// TIA Portal V21 program export: 0 tag tables, 0 data types, 1 data blocks, 1 code blocks (in call order from the OBs), 0 instance data blocks

DATA_BLOCK "DB_FAT_Demo"   // DB1
{ S7_Optimized_Access := 'FALSE' }
VERSION : 1.0
// SPDX-License-Identifier: MIT. Public passive laboratory example.
// stored: AutoNumber true, CodeModifiedDate 2026-11-03T19:44:32.7091278Z, CompileDate 2026-11-03T19:44:33.4739621Z, CreationDate 2026-11-03T19:44:31.2051572Z, DBAccessibleFromOPCUA true, DBAccessibleFromWebserver true, DownloadDate 0001-01-01T00:00:00Z, InterfaceModifiedDate 2026-11-03T19:44:32.7091278Z, IsConsistent true, IsKnowHowProtected false, IsOnlyStoredInLoadMemory false, IsPLCDB false, IsWriteProtectedInAS false, LoadMemoryLength 5286, ModifiedDate 2026-11-03T19:44:32.7091278Z, ParameterModified 2026-11-03T19:44:32.7091278Z, StructureModified 2026-11-03T19:44:32.7091278Z, WorkMemoryLength 192
   VAR RETAIN
      EnableDemo { ExternalAccessible := 'False'; ExternalVisible := 'False'; ExternalWritable := 'False'} : Bool := TRUE;   // isolated virtual copy only
      StopHealthy : Bool := TRUE;
      P101_Request : Bool := FALSE;
      P101_RequestedSpeed : Real := REAL#60.0;
      P101_RunCommand { ExternalWritable := 'False'} : Bool := FALSE;
      P101_SpeedCommand { ExternalWritable := 'False'} : Real := REAL#0.0;
      P101_Running : Bool := FALSE;
      P101_SpeedFeedback : Real := REAL#0.0;
      P101_Fault : Bool := FALSE;
      P201_Request : Bool := FALSE;
      P201_RequestedSpeed : Real := REAL#60.0;
      P201_RunCommand { ExternalWritable := 'False'} : Bool := FALSE;
      P201_SpeedCommand { ExternalWritable := 'False'} : Real := REAL#0.0;
      P201_Running : Bool := FALSE;
      P201_SpeedFeedback : Real := REAL#0.0;
      P201_Fault : Bool := FALSE;
      P202_Request : Bool := FALSE;
      P202_RequestedSpeed : Real := REAL#60.0;
      P202_RunCommand { ExternalWritable := 'False'} : Bool := FALSE;
      P202_SpeedCommand { ExternalWritable := 'False'} : Real := REAL#0.0;
      P202_Running : Bool := FALSE;
      P202_SpeedFeedback : Real := REAL#0.0;
      P202_Fault : Bool := FALSE;
      P301_Request : Bool := FALSE;
      P301_RequestedSpeed : Real := REAL#60.0;
      P301_RunCommand { ExternalWritable := 'False'} : Bool := FALSE;
      P301_SpeedCommand { ExternalWritable := 'False'} : Real := REAL#0.0;
      P301_Running : Bool := FALSE;
      P301_SpeedFeedback : Real := REAL#0.0;
      P301_Fault : Bool := FALSE;
      XV101_Request : Bool := FALSE;
      XV101_OpenCommand { ExternalWritable := 'False'} : Bool := FALSE;
      XV101_Open : Bool := FALSE;
      XV101_Closed : Bool := TRUE;
      XV201_Request : Bool := FALSE;
      XV201_OpenCommand { ExternalWritable := 'False'} : Bool := FALSE;
      XV201_Open : Bool := FALSE;
      XV201_Closed : Bool := TRUE;
      XV202_Request : Bool := FALSE;
      XV202_OpenCommand { ExternalWritable := 'False'} : Bool := FALSE;
      XV202_Open : Bool := FALSE;
      XV202_Closed : Bool := TRUE;
      XV301_Request : Bool := FALSE;
      XV301_OpenCommand { ExternalWritable := 'False'} : Bool := FALSE;
      XV301_Open : Bool := FALSE;
      XV301_Closed : Bool := TRUE;
      XV102_Request : Bool := FALSE;
      XV102_OpenCommand { ExternalWritable := 'False'} : Bool := FALSE;
      XV102_Open : Bool := FALSE;
      XV102_Closed : Bool := TRUE;
      XV203_Request : Bool := FALSE;
      XV203_OpenCommand { ExternalWritable := 'False'} : Bool := FALSE;
      XV203_Open : Bool := FALSE;
      XV203_Closed : Bool := TRUE;
      XV103_Request : Bool := FALSE;
      XV103_OpenCommand { ExternalWritable := 'False'} : Bool := FALSE;
      XV103_Open : Bool := FALSE;
      XV103_Closed : Bool := TRUE;
      FCV302_RequestedPosition : Real := REAL#0.0;
      FCV302_PositionCommand { ExternalWritable := 'False'} : Real := REAL#0.0;
      FCV302_PositionFeedback : Real := REAL#0.0;
      LT101_Raw : Int := INT#16589;
      LT101_Percent { ExternalWritable := 'False'} : Real := REAL#0.0;
      TK101_Volume : Real := REAL#720.0;
      LSL101 : Bool := FALSE;
      LSH101 : Bool := FALSE;
      LT201_Raw : Int := INT#6912;
      LT201_Percent { ExternalWritable := 'False'} : Real := REAL#0.0;
      TK201_Volume : Real := REAL#450.0;
      LSL201 : Bool := FALSE;
      LSH201 : Bool := FALSE;
      LT301_Raw : Int := INT#4147;
      LT301_Percent { ExternalWritable := 'False'} : Real := REAL#0.0;
      TK301_Volume : Real := REAL#180.0;
      LSL301 : Bool := FALSE;
      LSH301 : Bool := FALSE;
   END_VAR
BEGIN
END_DATA_BLOCK

ORGANIZATION_BLOCK "Main"   // OB1, SCL, ProgramCycle
{ S7_Optimized_Access := 'TRUE' }
VERSION : 1.0
// SPDX-License-Identifier: MIT. No equipment library or process sequence.
// stored: AutoNumber true, CodeModifiedDate 2026-11-03T19:44:43.8400479Z, CompileDate 2026-11-03T19:44:43.8400479Z, ConstantName OB_Main, CreationDate 2026-11-03T19:44:33.7000652Z, DownloadDate 0001-01-01T00:00:00Z, EventClass Program cycle, HandleErrorsWithinBlock false, InterfaceModifiedDate 2026-11-03T19:44:33.988557Z, IsConsistent true, IsIECCheckEnabled false, IsKnowHowProtected false, IsWriteProtected false, LoadMemoryLength 14729, ModifiedDate 2026-11-03T19:44:43.8400479Z, PLCSimAdvancedSupport true, ParameterModified 2026-11-03T19:44:33.9885569Z, PriorityNumber 1, ProcessImagePartNumber 65535, SetENOAutomatically false, StructureModified 2026-11-03T19:44:33.988557Z, VirtualPlcSupport false, WorkMemoryLength 554
   VAR_INPUT
      Initial_Call : Bool;   // Initial call of this OB
      Remanence : Bool;   // =True, if remanent data are available
   END_VAR
BEGIN

       "DB_FAT_Demo".P101_RunCommand := "DB_FAT_Demo".EnableDemo AND "DB_FAT_Demo".StopHealthy AND "DB_FAT_Demo".P101_Request;
       IF "DB_FAT_Demo".P101_RunCommand THEN
           "DB_FAT_Demo".P101_SpeedCommand := LIMIT(MN := REAL#0.0, IN := "DB_FAT_Demo".P101_RequestedSpeed, MX := REAL#100.0);
       ELSE
           "DB_FAT_Demo".P101_SpeedCommand := REAL#0.0;
       END_IF;
       "DB_FAT_Demo".P201_RunCommand := "DB_FAT_Demo".EnableDemo AND "DB_FAT_Demo".StopHealthy AND "DB_FAT_Demo".P201_Request;
       IF "DB_FAT_Demo".P201_RunCommand THEN
           "DB_FAT_Demo".P201_SpeedCommand := LIMIT(MN := REAL#0.0, IN := "DB_FAT_Demo".P201_RequestedSpeed, MX := REAL#100.0);
       ELSE
           "DB_FAT_Demo".P201_SpeedCommand := REAL#0.0;
       END_IF;
       "DB_FAT_Demo".P202_RunCommand := "DB_FAT_Demo".EnableDemo AND "DB_FAT_Demo".StopHealthy AND "DB_FAT_Demo".P202_Request;
       IF "DB_FAT_Demo".P202_RunCommand THEN
           "DB_FAT_Demo".P202_SpeedCommand := LIMIT(MN := REAL#0.0, IN := "DB_FAT_Demo".P202_RequestedSpeed, MX := REAL#100.0);
       ELSE
           "DB_FAT_Demo".P202_SpeedCommand := REAL#0.0;
       END_IF;
       "DB_FAT_Demo".P301_RunCommand := "DB_FAT_Demo".EnableDemo AND "DB_FAT_Demo".StopHealthy AND "DB_FAT_Demo".P301_Request;
       IF "DB_FAT_Demo".P301_RunCommand THEN
           "DB_FAT_Demo".P301_SpeedCommand := LIMIT(MN := REAL#0.0, IN := "DB_FAT_Demo".P301_RequestedSpeed, MX := REAL#100.0);
       ELSE
           "DB_FAT_Demo".P301_SpeedCommand := REAL#0.0;
       END_IF;
       "DB_FAT_Demo".XV101_OpenCommand := "DB_FAT_Demo".EnableDemo AND "DB_FAT_Demo".StopHealthy AND "DB_FAT_Demo".XV101_Request;
       "DB_FAT_Demo".XV201_OpenCommand := "DB_FAT_Demo".EnableDemo AND "DB_FAT_Demo".StopHealthy AND "DB_FAT_Demo".XV201_Request;
       "DB_FAT_Demo".XV202_OpenCommand := "DB_FAT_Demo".EnableDemo AND "DB_FAT_Demo".StopHealthy AND "DB_FAT_Demo".XV202_Request;
       "DB_FAT_Demo".XV301_OpenCommand := "DB_FAT_Demo".EnableDemo AND "DB_FAT_Demo".StopHealthy AND "DB_FAT_Demo".XV301_Request;
       "DB_FAT_Demo".XV102_OpenCommand := "DB_FAT_Demo".EnableDemo AND "DB_FAT_Demo".StopHealthy AND "DB_FAT_Demo".XV102_Request;
       "DB_FAT_Demo".XV203_OpenCommand := "DB_FAT_Demo".EnableDemo AND "DB_FAT_Demo".StopHealthy AND "DB_FAT_Demo".XV203_Request;
       "DB_FAT_Demo".XV103_OpenCommand := "DB_FAT_Demo".EnableDemo AND "DB_FAT_Demo".StopHealthy AND "DB_FAT_Demo".XV103_Request;
       IF "DB_FAT_Demo".EnableDemo AND "DB_FAT_Demo".StopHealthy THEN
           "DB_FAT_Demo".FCV302_PositionCommand := LIMIT(MN := REAL#0.0, IN := "DB_FAT_Demo".FCV302_RequestedPosition, MX := REAL#100.0);
       ELSE
           "DB_FAT_Demo".FCV302_PositionCommand := REAL#0.0;
       END_IF;
       "DB_FAT_Demo".LT101_Percent := SCALE_X(MIN := REAL#0.0,
           VALUE := NORM_X(MIN := INT#0, VALUE := "DB_FAT_Demo".LT101_Raw, MAX := INT#27648), MAX := REAL#100.0);
       "DB_FAT_Demo".LT201_Percent := SCALE_X(MIN := REAL#0.0,
           VALUE := NORM_X(MIN := INT#0, VALUE := "DB_FAT_Demo".LT201_Raw, MAX := INT#27648), MAX := REAL#100.0);
       "DB_FAT_Demo".LT301_Percent := SCALE_X(MIN := REAL#0.0,
           VALUE := NORM_X(MIN := INT#0, VALUE := "DB_FAT_Demo".LT301_Raw, MAX := INT#27648), MAX := REAL#100.0);
END_ORGANIZATION_BLOCK
